Staubli VAL3: saveLog.pgx

public program saveLog(string x_sPath (dimensions=1), num& x_nResult (dimensions=1))
  local num l_n
  local num l_nLogMsgIndex
begin
  if x_sPath==""
    x_nResult=Log:libSave()
  else
    x_nResult=Log:libSave(x_sPath)
  endIf
  delay(0.5)
end
